(* IEC 61131-3 sources: PortalRobot/Portal_robot/Device/application/ST/ST_MOTION_MANAGER, 7 files *)

(* ---- E_MOTION_MANAGER_STATE.st ---- *)
{attribute 'qualified_only'}
{attribute 'strict'}
TYPE E_MOTION_MANAGER_STATE :
(
	IDLE,
	VALIDATE,
	MOTION_SIM,
	MOTION_MODBUS,
	DONE,
	ERROR
);
END_TYPE

(* ---- ST_MOTION_MANAGER.st ---- *)
TYPE ST_MOTION_MANAGER :
STRUCT
	Command : ST_MOTION_MANAGER_COMMAND; // Команды менеджеру движения
	Status  : ST_MOTION_MANAGER_STATUS; // Рабочие статусы менеджера движения
	Diag    : ST_MOTION_MANAGER_DIAG; // Состояние автомата менеджера движения
	Error   : ST_MOTION_MANAGER_ERRORS; // Активные и последние ошибки
END_STRUCT
END_TYPE

(* ---- ST_MOTION_MANAGER_COMMAND.st ---- *)
TYPE ST_MOTION_MANAGER_COMMAND :
STRUCT
	eTargetPoint : E_POINT_NAME; // Имя целевой точки
	xGlobalError : BOOL; // Глобальная ошибка ячейки
	xExecute     : BOOL; // Команда запуска движения
	xStop        : BOOL; // Штатная операторская остановка без формирования аварии
	xReset       : BOOL; // Команда сброса ошибки
	xMode        : BOOL; // TRUE: Modbus, FALSE: SoftMotion
END_STRUCT
END_TYPE

(* ---- ST_MOTION_MANAGER_DIAG.st ---- *)
TYPE ST_MOTION_MANAGER_DIAG :
STRUCT
	eState : E_MOTION_MANAGER_STATE; // Текущее состояние автомата движения
	stWarning : ST_WARNING_EVENT; // Последнее предупреждение менеджера движения
END_STRUCT
END_TYPE

(* ---- ST_MOTION_MANAGER_ERROR.st ---- *)
TYPE ST_MOTION_MANAGER_ERROR :
STRUCT
	POINT_INVALID : BOOL; // Целевая точка не прошла проверку
	GROUP_ERROR   : BOOL; // Группа осей завершила движение с ошибкой
	GLOBAL_STOP   : BOOL; // Получена глобальная ошибка ячейки
	START_TIMEOUT : BOOL; // Истекло ожидание проверки точки или старта группы
END_STRUCT
END_TYPE

(* ---- ST_MOTION_MANAGER_ERRORS.st ---- *)
TYPE ST_MOTION_MANAGER_ERRORS :
STRUCT
	dwErrorActive : DWORD; // Битовая маска активных ошибок
	dwErrorLast   : DWORD; // Битовая маска последних ошибок
	dwAlarmActive : DWORD; // Собственные аварии менеджера движения для общего журнала
	stErrorActive : ST_MOTION_MANAGER_ERROR; // Расшифровка активных ошибок
	stErrorLast   : ST_MOTION_MANAGER_ERROR; // Расшифровка последних ошибок
END_STRUCT
END_TYPE

(* ---- ST_MOTION_MANAGER_STATUS.st ---- *)
TYPE ST_MOTION_MANAGER_STATUS :
STRUCT
	xReady        : BOOL; // Менеджер готов принять команду
	xBusy         : BOOL; // Выполняется движение
	xDone         : BOOL; // Движение завершено
	xError        : BOOL; // Менеджер находится в ошибке
	eCurrentPoint : E_POINT_NAME; // Последняя достигнутая точка
END_STRUCT
END_TYPE
